(* IEC 61131-3 sources: JingjiangArm/moonboxpro_arm_8.4/Application/Application/任务列表/TensionTask/电机运动/MotionCtl_Gear/PrnVelCtl, 9 files *)

(* ---- KS_CalcMovePara.st ---- *)
(*@CES
Name=KS_CalcMovePara
Type=FunctionBlock
TypeGuid=6f9dac99-8de1-4efc-8465-68ac443b7d08
Guid=11217540-9eff-4725-bda6-b930b9e4eccf
HasDeclaration=True
HasImplementation=True
*)
{DECLARATION}
FUNCTION KS_CalcMovePara : LREAL(*计算运动时间参数|
								控制为even段|只考虑了目标轴匀速、当前轴加速
								返回值作为最终的加速时间s|
								如果时间不能被运动时间间隔整除则会存在pt写入按照整数个
								时间间隔，这里监控的p是使用实际时间的，但是对最终的位置偏差
								没影响。
								负值为返回错误
								-1 参数错误*)
VAR_INPUT
	i_lrVelSa:LREAL;(*启动速度m/min|V0*)
	i_lrVelTar:LREAL;(*目标速度m/min|Vt*)
	i_iDeltime:INT:=21;(*速度规划间隔时间ms|pt运动时间*)
	i_lrGirth_Axis:LREAL;(*轴周长|mm*)
	i_lrReductionRatio:LREAL;(*减速比|电机侧/版辊侧*)
	i_lrDeltPos_Init:LREAL;(*初始位置偏差Pul|开始运动时目标轴和当前轴的位置p偏差*)
	i_lrDeltPos_Final:LREAL;(*最终偏差Pul|最终的目标轴和当前轴的p偏差*)
	i_dwMotorPPR:DWORD:=2097152;(*电机运动一圈的值*)
	i_iSetTime:INT;(*用来计算模数s|*)
END_VAR
VAR
	lrDeltV: LREAL;(*mm/ms*)
	uiTime_N: UINT;(**)
	iDeltT: INT;(*ms*)
	lrCoeff_Axis: LREAL;(*当前轴的比例|Pul/mm*)
	lrRtnValue: LREAL:=0;(*返回值*)
	lrVt: LREAL;(*mm/ms*)
	lrVo: LREAL;(*mm/ms*)
	lrGirth_Axis: LREAL;
	lrDeltPos_Init: LREAL;(*Pul*)
	lrDeltPos_Final:LREAL;(*Pul*)
	(*计算临时变量*)
	uiModCoeff: UINT;(*圈数取整值*)

	lrTemp: LREAL;
	lrTemp1: LREAL;

	(*目标轴位移|mm*)
	lrS_Tar: LREAL;
	(*当前轴位移|mm*)
	lrS_Cur: LREAL;
	dwTime_ms:DWORD;
	lrDelP: LREAL;
	lrDeltS: LREAL;
	lrTime:LREAL;

	lrWatchS_Tar: LREAL;
	lrWatchS_Cur: LREAL;
	lrWatchP_Tar: LREAL;
	lrWatchP_Cur: LREAL;
	lrA: LREAL;
	uiN: UINT;
	iSetTime: INT;
END_VAR
{IMPLEMENTATION}
IF i_lrVelTar<=i_lrVelSa THEN
	lrRtnValue:=-1;
END_IF
lrVt:=i_lrVelTar/60;
lrVo:=i_lrVelSa/60;
lrDeltV:=lrVt-lrVo;

iDeltT:=i_iDeltime;
IF i_iDeltime<=0 THEN
	lrRtnValue:=-1;
END_IF

(*当前轴周长*)
lrGirth_Axis:=i_lrGirth_Axis;
IF lrGirth_Axis<=0 THEN
	lrRtnValue:=-1;
END_IF

IF i_dwMotorPPR<=0 THEN
	lrRtnValue:=-1;
END_IF

IF i_lrReductionRatio<=0 THEN
	lrRtnValue:=-1;
END_IF

(*初始位置偏差Pul|开始运动时目标轴和当前轴的位置p偏差*)
lrDeltPos_Init:=i_lrDeltPos_Init;
lrDeltPos_Init:=KS_MOD_LREAL(lrDeltPos_Init,(i_dwMotorPPR*i_lrReductionRatio));

(*最终偏差Pul|最终的目标轴和当前轴的p偏差*)
lrDeltPos_Final:=i_lrDeltPos_Final;
lrDeltPos_Final:=KS_MOD_LREAL(lrDeltPos_Final,(i_dwMotorPPR*i_lrReductionRatio));

iSetTime:=i_iSetTime;
IF i_iSetTime>=500 THEN(*防止溢出*)
	iSetTime:=500;
END_IF

IF lrRtnValue=0 THEN(*未有错误*)
	dwTime_ms:=(iSetTime)*1000;
	uiTime_N:=(iSetTime)*1000/iDeltT;
	lrA:=lrDeltV/dwTime_ms;

	(*当前轴比例|版辊距离mm转换为电机脉冲值*)
	lrCoeff_Axis:=i_lrReductionRatio*i_dwMotorPPR/i_lrGirth_Axis;(*Pul/mm*)

	(*计算模数值*)
	(*运动的位移*)
	lrS_Tar:=lrVt*dwTime_ms;(*mm*)
	lrS_Cur:=uiTime_N*lrVo*iDeltT+0.5*lrA*iDeltT*iDeltT*uiTime_N*(1+uiTime_N)+
			lrVt*(dwTime_ms-uiTime_N*iDeltT);(*mm*)
	lrDeltS:=lrS_Tar-lrS_Cur;
	IF lrDeltS<=0 THEN
		lrRtnValue:=-2;
	END_IF

	(*转换为电机侧的脉冲*)
	lrDelP:=lrDeltS*lrCoeff_Axis;

	lrTemp:=lrDeltPos_Init+lrDelP-lrDeltPos_Final;
	IF lrTemp<=0 THEN
		lrRtnValue:=-3;
	END_IF
	lrTemp1:=i_dwMotorPPR*i_lrReductionRatio;

	lrTemp:=lrTemp/lrTemp1;
	(*取整数*)

	(*圈数值取整数|版辊圈数*)
	uiModCoeff:=LREAL_TO_UINT(lrTemp);
	IF uiModCoeff<lrTemp THEN
		uiModCoeff:=uiModCoeff+1;
	END_IF

	(*计算需要的时间|按照这个时间可以在目标速度时达到位置同步*)
	IF lrRtnValue=0 THEN
		(*反算时间*)
		lrDelP:=lrDeltPos_Final+uiModCoeff*i_lrReductionRatio*i_dwMotorPPR-lrDeltPos_Init;
		lrDeltS:=lrDelP/lrCoeff_Axis;

		(*寻找复合条件的时间|时间/21的余数小于21*)
		FOR uiN:=uiTime_N TO uiTime_N+10000  BY 1 DO
			lrTemp:=lrDeltV*iDeltT*iDeltT*(1+uiN)*uiN*0.5;
			lrTemp1:=(-lrDeltS-uiN*lrVo*iDeltT+uiN*iDeltT*lrVt);
			lrTime:=lrTemp/lrTemp1;

			IF lrTime-uiN*iDeltT<=iDeltT THEN
				EXIT;
			END_IF

			IF uiN=uiTime_N+10000 THEN(*没有找到|输出负值 标记*)
				lrTime:=-4;
			END_IF
		END_FOR

	END_IF

	IF lrRtnValue=0 THEN
		lrRtnValue:=LREAL_TO_REAL(lrTime/1000);

		(*用于监控*)
		lrWatchS_Tar:=lrVt*lrTime;(*mm*)
		uiTime_N:=uiN;
		lrA:=lrDeltV/lrTime;
		lrWatchS_Cur:=uiTime_N*lrVo*iDeltT+0.5*lrA*iDeltT*iDeltT*uiTime_N*(1+uiTime_N)+
					lrVt*(lrTime-uiTime_N*iDeltT);(*mm*)
		lrWatchP_Tar:=lrWatchS_Tar*lrCoeff_Axis;
		lrWatchP_Cur:=lrWatchS_Cur*lrCoeff_Axis;
	END_IF
END_IF
KS_CalcMovePara:=lrRtnValue;

(* ---- KS_GetInitSts.st ---- *)
(*@CES
Name=KS_GetInitSts
Type=FunctionBlock
TypeGuid=6f9dac99-8de1-4efc-8465-68ac443b7d08
Guid=7ae6f696-fe0b-48ae-942d-bfb0aac909fe
HasDeclaration=True
HasImplementation=True
*)
{DECLARATION}
FUNCTION KS_GetInitSts : BYTE(*获取初始值状态|返回修改的状态*)
VAR_INPUT
	i_bySwitchType:BYTE;(*切换方式|0-空转状态下不考虑单联动状态下都可以切换运动状态
								  |1-空转状态下只有处于联动状态下的轴可以切换*)
	i_xLinkageKnob: BOOL;(*联动旋钮*)
	i_xLinkageSts: BOOL;(*联动状态*)
END_VAR
VAR
	byAxisMotionSts: BYTE;
END_VAR
{IMPLEMENTATION}
IF i_bySwitchType=0 THEN(*空转状态下不考虑单联动状态下都可以切换运动状态*)
	IF i_xLinkageKnob THEN
		byAxisMotionSts:= 0;
	ELSE
		byAxisMotionSts:= 2;
	END_IF
ELSIF i_bySwitchType=1 THEN(*空转状态下只有处于联动状态下的轴可以切换*)
	IF i_xLinkageSts THEN
		byAxisMotionSts:=0;
	ELSE
		byAxisMotionSts:=2;
	END_IF
END_IF
KS_GetInitSts:=byAxisMotionSts;

(* ---- KS_GetMotionSts.st ---- *)
(*@CES
Name=KS_GetMotionSts
Type=FunctionBlock
TypeGuid=6f9dac99-8de1-4efc-8465-68ac443b7d08
Guid=c01ac71d-e678-459d-bed7-b9a659b9ae68
HasDeclaration=True
HasImplementation=True
*)
{DECLARATION}
FUNCTION KS_GetMotionSts : BOOL(*色组轴的运动状态处理|只在开机时候使用 同时控制压辊合压状态|Liu.yt
										轴运动状态标志|0:同步运动状态.
													  |1:同步运动时停止运动状态.
													  |2:停止运动状态
													  |3:停止运动时加速到单运行速度状态.
													  |4:单运行时减速到停止状态.
													  |5:停止运动时或者使用单运行速度运行时加速到同步运动状态.
													  |6:非同步运动时急停到0状态.
													  |7:非同步运动时空转停机到0状态.*)
(*2022.9.21.154927 6,7步中停止的条件判断写错了*)
(*2022.11.29.232720 轴速度是带方向|作为条件需要增加取绝对值*)
(*2023.11.27.165212 增加印刷是否能切换单联动的选择输入接口*)
VAR_INPUT
	i_iGrpId: INT;
	i_xMotionStsSwitchEn:BOOL;(*切换使能|使用该功能需要常有效*)
	i_bySwitchType:BYTE;(*切换方式|0-空转状态下不考虑单联动状态下都可以切换运动状态
								  |1-空转状态下只有处于联动状态下的轴可以切换*)
	i_iGrpAxisNum_Pu: INT; (*色组轴数量*)
	i_pstStSysParam: POINTER TO StSysParam;
//	i_pstStGrpParam: POINTER TO StGrpParam;(*系参数访问入口|*)
	i_paiGrpAxisList: POINTER TO ARRAY [1..MAX_STATION_NUM] OF INT; (*系内所有轴的列表*)
//	i_pastStAxisParam: POINTER TO ARRAY [1..MAX_STATION_NUM] OF StAxisParam;
	i_pastStIOMap_Main_FE						: POINTER TO ARRAY [1..4] OF StIOMap_Main_FE;(*轴io数据区域|AB系*)
	i_pastStIOMap_Axis_FE					: POINTER TO ARRAY [1..MAX_UNIT_NUM] OF StIOMap_Axis_FE;(*轴io数据区域|`````````````````````````````````````````````*)
//	i_pastStIOMap_AxisBasic: POINTER TO ARRAY [1..MAX_STATION_NUM] OF StIOMap_AxisBasic;(*基础io映射表|*)
	i_pabyAxisMotionSts: POINTER TO ARRAY [1..MAX_STATION_NUM] OF BYTE;(*轴运动状态|*)
	i_paxAxisInching:POINTER TO ARRAY [1..MAX_STATION_NUM] OF BOOL;(*轴在单运行|用于控制单运行指示灯显示*)
	i_paxLastAxisInchBtn:POINTER TO ARRAY [1..MAX_STATION_NUM] OF BOOL;(*轴的单运行按钮保留值|用于判断沿*)
	i_iMaxVel_StsSwitch:INT;(*状态切换的最大速度*)
	i_pxFlag_StsSwitchEn:POINTER TO BOOL;(*状态切换使能标志@内部的状态切换标志*)
	i_xChangLinkageStsWhenPrint:BOOL;(*印刷时候可以切换单联动@2023.11.27.164606*)
END_VAR
VAR

	iN: INT;
	xFlag_StsSwitchEn: BOOL;(*状态切换标志*)
	xStsSwitchEn: BOOL;(*状态切换使能*)
	xRetainStsEn: BOOL;(*保持状态标志*)
	iUnitId: INT;
	byAxisMotionSts: BYTE;
	xLastAxisInchBtn: BOOL;
	xAxisInching: BOOL;
	pstStUnitParam_Save: POINTER TO StUnitParam_Save;
	pstStUnitParam_UnSave: POINTER TO StUnitParam_UnSave;
	pstStGrpParam_Save: POINTER TO StGrpParam_Save;
	pstStGrpParam_UnSave: POINTER TO StGrpParam_UnSave;
	pstStIOMap_Axis_FE: POINTER TO StIOMap_Axis_FE;
	xCanSwitchSts_CurAxis: BOOL;(*当前轴可以切换状态标志*)
	dwAxisMotionStsNotOk: DWORD;
END_VAR
{IMPLEMENTATION}
IF i_pstStSysParam<>0 AND
	i_paiGrpAxisList<>0 AND
	i_pastStIOMap_Main_FE<>0 AND
	i_pastStIOMap_Axis_FE<>0 AND
	i_pabyAxisMotionSts<>0 AND
	i_paxAxisInching<>0 AND
	i_paxLastAxisInchBtn<>0 AND
	i_iGrpAxisNum_Pu>0 AND
	i_pxFlag_StsSwitchEn<>0 THEN(*参数合法*)

	xFlag_StsSwitchEn:=i_pxFlag_StsSwitchEn^;
	pstStGrpParam_Save:= ADR(i_pstStSysParam^.astStGrpParam_Save[i_iGrpId]);
	pstStGrpParam_UnSave:= ADR(i_pstStSysParam^.astStGrpParam_UnSave[i_iGrpId]);
	(*2023.11.27.171042 增加了印刷时候有单联动切换的选择接口*)
	xStsSwitchEn:= (pstStGrpParam_UnSave^.xFlag_Ink OR(*空转状态下可以使用|*)
					(pstStGrpParam_UnSave^.xFlag_Print AND i_xChangLinkageStsWhenPrint)) AND
					pstStGrpParam_UnSave^.rVel_Cur<=i_iMaxVel_StsSwitch;(*小于速度限制可以使用*)
	(*印刷时候或者超过限制速度时候|与xStsSwitchEn搭配使用*)
	xRetainStsEn:=(pstStGrpParam_UnSave^.xFlag_Print AND NOT i_xChangLinkageStsWhenPrint)
				OR pstStGrpParam_UnSave^.rVel_Cur>i_iMaxVel_StsSwitch;

	(*切换条件处理*)
	IF  xStsSwitchEn THEN
		xFlag_StsSwitchEn:=TRUE;
	END_IF

	IF i_xMotionStsSwitchEn THEN
		FOR iN:=1 TO i_iGrpAxisNum_Pu BY 1 DO
			iUnitId:=i_paiGrpAxisList^[iN];
			pstStUnitParam_Save:=ADR(i_pstStSysParam^.astStUnitParam_Save[iUnitId]);
			pstStUnitParam_UnSave:=ADR(i_pstStSysParam^.astStUnitParam_UnSave[iUnitId]);
			pstStIOMap_Axis_FE:=ADR(i_pastStIOMap_Axis_FE^[iUnitId]);
			byAxisMotionSts:=i_pabyAxisMotionSts^[iUnitId];
			xLastAxisInchBtn:=i_paxLastAxisInchBtn^[iUnitId];
			xAxisInching:=i_paxAxisInching^[iUnitId];

			xCanSwitchSts_CurAxis:=FALSE;
			IF i_bySwitchType=0 THEN(*空转状态下不考虑单联动状态下都可以切换运动状态*)
				xCanSwitchSts_CurAxis:= pstStUnitParam_UnSave^.xMoveEnable_Motor;
			ELSIF i_bySwitchType=1 THEN(*空转状态下只有处于联动状态下的轴可以切换*)
				xCanSwitchSts_CurAxis:= pstStUnitParam_Save^.xLinkage;
			END_IF

			IF xCanSwitchSts_CurAxis THEN
				CASE byAxisMotionSts OF
					0:(*同步运动状态|此时检查但联动旋钮的状态*)
						IF NOT pstStIOMap_Axis_FE^.i_xLinkage AND (*切换到单动状态*)
							NOT pstStIOMap_Axis_FE^.o_xRel_Press THEN(*压辊未合压时起作用*)
							byAxisMotionSts:=1;
						END_IF
					1:(*处于停止运动过程状态|等待到达停止运动状态*)
						IF pstStIOMap_Axis_FE^.i_xLinkage THEN(*联动状态|恢复到同步运动状态*)
							byAxisMotionSts:=5;
						END_IF

						IF byAxisMotionSts=1 THEN
							IF ABS(pstStUnitParam_UnSave^.rAxisVel_PrnRoller)<=0.0001 THEN(*减速到0我们认为到达了停止运动状态*)
								byAxisMotionSts:=2;
							END_IF
						END_IF
					2:(*停止运动状态*)
						IF pstStIOMap_Axis_FE^.i_xLinkage THEN(*联动状态|恢复到同步运动状态*)
							byAxisMotionSts:=5;
						END_IF

						(*检查单运行是否按下*)
						IF byAxisMotionSts=2 THEN
							IF pstStIOMap_Axis_FE^.i_xInch AND NOT xLastAxisInchBtn THEN(*单运行按下了*)
								byAxisMotionSts:=3;
							END_IF
						END_IF

					3:(*加速到单运行状态*)
						IF pstStIOMap_Axis_FE^.i_xLinkage THEN(*联动状态|恢复到同步运动状态*)
							byAxisMotionSts:=5;
						END_IF

						IF byAxisMotionSts=3 THEN
							IF (pstStIOMap_Axis_FE^.i_xInch AND NOT xLastAxisInchBtn) OR(*单运行按下了*)
								NOT xStsSwitchEn THEN(*退出了状态*)
								byAxisMotionSts:=4;
							END_IF
						END_IF
					4:(*单运行状态停止到停止状态*)
						IF pstStIOMap_Axis_FE^.i_xLinkage THEN(*联动状态|恢复到同步运动状态*)
							byAxisMotionSts:=5;
						END_IF

						IF byAxisMotionSts=4 THEN
							IF ABS(pstStUnitParam_UnSave^.rAxisVel_PrnRoller)<=0.0001 THEN(*减速到0我们认为到达了停止运动状态*)
								byAxisMotionSts:=2;
							END_IF
						END_IF
					5:(*前往同步运动状态*)
						IF NOT pstStIOMap_Axis_FE^.i_xLinkage THEN(*切换到单动状态*)
							byAxisMotionSts:=1;
						END_IF

						IF byAxisMotionSts=5 THEN
							IF ABS(ABS(pstStUnitParam_UnSave^.rAxisVel_PrnRoller)-pstStGrpParam_UnSave^.rVel_Cur)<=0.0001 THEN(*到达当前速度*)
								byAxisMotionSts:=0;
							END_IF
						END_IF
					6,7:(*非同步状态下非停止状态下的停止和急停*)
						IF ABS(pstStUnitParam_UnSave^.rAxisVel_PrnRoller)<=0.0001 THEN(*到达0速度|2022.9.21.154723 -以前的条件写错了*)
							byAxisMotionSts:=KS_GetInitSts(i_bySwitchType,
													pstStIOMap_Axis_FE^.i_xLinkage,
													pstStUnitParam_Save^.xLinkage);
						END_IF
				ELSE
					byAxisMotionSts:=KS_GetInitSts(i_bySwitchType,
											pstStIOMap_Axis_FE^.i_xLinkage,
											pstStUnitParam_Save^.xLinkage);
				END_CASE
			ELSE
				byAxisMotionSts:=KS_GetInitSts(i_bySwitchType,
										pstStIOMap_Axis_FE^.i_xLinkage,
										pstStUnitParam_Save^.xLinkage);
			END_IF

			(*处理单运行指示*)
			IF byAxisMotionSts=3 OR(*单运行加速*)
				byAxisMotionSts=4 THEN(*单运行减速*)
				xAxisInching:=TRUE;
			ELSE
				xAxisInching:=FALSE;
			END_IF

			(*切换使能无效了-在状态恢复到初始状态时候xFlag_StsSwitchEn标志为false|
			byAxisMotionSts 在停机时候强制写为初值|
							在印刷状态或者超过限制速度时不切换|*)
			IF xRetainStsEn THEN(*保持之前状态|*)
				byAxisMotionSts:=i_pabyAxisMotionSts^[iUnitId];
			ELSE
				IF NOT xFlag_StsSwitchEn THEN
					byAxisMotionSts:=KS_GetInitSts(i_bySwitchType,
												pstStIOMap_Axis_FE^.i_xLinkage,
												pstStUnitParam_Save^.xLinkage);
				END_IF
			END_IF

			(*处理停机和急停*)
			IF byAxisMotionSts<>0 AND  byAxisMotionSts<>2 THEN
				IF pstStGrpParam_UnSave^.xFlag_EStoping THEN(*急停过程中|*)
					byAxisMotionSts:=6;
				ELSIF pstStGrpParam_UnSave^.xFlag_Ink AND
					(pstStGrpParam_UnSave^.xFlag_Stoping OR (*空转停止过程中*)
					pstStGrpParam_UnSave^.xFlag_FastStoping) THEN
					byAxisMotionSts:=7;
				END_IF

				(*判断轴运动状态|未处于停止状态或者同步状态|*)
				dwAxisMotionStsNotOk:=dwAxisMotionStsNotOk OR SHL(DWORD#1,iUnitId-1);
			END_IF

			(*使能模式控制|2022.7.14.121739*)
			IF i_bySwitchType=0 THEN
				IF byAxisMotionSts=2 THEN(*停止状态 写3*)
					pstStUnitParam_Save^.wEnableMode_Motor:=3;
				ELSE(*非停止状态|写4*)
					pstStUnitParam_Save^.wEnableMode_Motor:=4;
				END_IF
			ELSE
				IF pstStUnitParam_Save^.wEnableMode_Motor=3 OR
					pstStUnitParam_Save^.wEnableMode_Motor=4 THEN(*说明进行过使能切换|此时强制将使能模式写成4*)
					pstStUnitParam_Save^.wEnableMode_Motor:=4;
				ELSE
					pstStUnitParam_Save^.wEnableMode_Motor:=0;
				END_IF
			END_IF

			i_pabyAxisMotionSts^[iUnitId]:=byAxisMotionSts;
			i_paxAxisInching^[iUnitId]:=xAxisInching;
			i_paxLastAxisInchBtn^[iUnitId]:=i_pastStIOMap_Axis_FE^[iUnitId].i_xInch;
		END_FOR

		(*切换条件处理*)
		IF NOT xStsSwitchEn THEN
			IF xFlag_StsSwitchEn THEN
				IF dwAxisMotionStsNotOk=0 THEN(*都处于初始态|可以清除标志了*)
					xFlag_StsSwitchEn:=FALSE;
				END_IF
			END_IF
		END_IF
	ELSE(*不使能*)
		FOR iN:=1 TO i_iGrpAxisNum_Pu BY 1 DO
			iUnitId:=i_paiGrpAxisList^[iN];
			pstStUnitParam_Save:=ADR(i_pstStSysParam^.astStUnitParam_Save[iUnitId]);
			pstStUnitParam_UnSave:=ADR(i_pstStSysParam^.astStUnitParam_UnSave[iUnitId]);
			i_pabyAxisMotionSts^[iUnitId]:=0;
			i_paxAxisInching^[iUnitId]:=FALSE;
			i_paxLastAxisInchBtn^[iUnitId]:=FALSE;

			IF pstStUnitParam_Save^.wEnableMode_Motor=3 OR
				pstStUnitParam_Save^.wEnableMode_Motor=4 THEN(*说明进行过使能切换|此时强制将使能模式写成4*)
				pstStUnitParam_Save^.wEnableMode_Motor:=4;
			ELSE
				pstStUnitParam_Save^.wEnableMode_Motor:=0;
			END_IF
		END_FOR
		xFlag_StsSwitchEn:=FALSE;
	END_IF

	i_pxFlag_StsSwitchEn^:=xFlag_StsSwitchEn;
END_IF

(* ---- KS_GetRelatePos.st ---- *)
(*@CES
Name=KS_GetRelatePos
Type=FunctionBlock
TypeGuid=6f9dac99-8de1-4efc-8465-68ac443b7d08
Guid=64bf2139-19b0-44f0-86e4-ed0fdab8fbfc
HasDeclaration=True
HasImplementation=True
*)
{DECLARATION}
FUNCTION KS_GetRelatePos : BOOL(*计算所有目标轴和当前轴的相对位置|节省空间就只做16个轴
								目标轴为联动非涂布轴*)
VAR_INPUT
	i_iAxisId_Cur:INT;(*当前轴id*)
	i_iGrpAxisNum_Pu: INT; (*色组轴数量*)
	i_paiGrpAxisList: POINTER TO ARRAY [1..MAX_UNIT_NUM] OF INT; (*系内所有轴的列表*)
	i_pastStUnitParam_Save: POINTER TO ARRAY [1..MAX_UNIT_NUM] OF StUnitParam_Save;
	i_pastStUnitParam_UnSave: POINTER TO ARRAY [1..MAX_UNIT_NUM] OF StUnitParam_UnSave;
	i_palrRelatePos:POINTER TO ARRAY [1..MAX_UNIT_NUM] OF LREAL;(*索引为目标轴*)
END_VAR
VAR
	in: INT;
	iAxisId: INT;
	pstStUnitParam_Save: POINTER TO StUnitParam_Save;
	pstStUnitParam_UnSave: POINTER TO StUnitParam_UnSave;
	pstStUnitParam_Cur_UnSave: POINTER TO StUnitParam_UnSave;
	ailist: ARRAY [1..MAX_STATION_NUM] OF INT;(*联动非涂布列表|不包含当前色*)
	iIndex:INT;
	xDne: BOOL;(*获取成功了*)
END_VAR
{IMPLEMENTATION}
(*初始化*)
IF	i_palrRelatePos<>0	THEN
	FOR iN:=1 TO 16 BY 1 DO
		i_palrRelatePos^[iN]:=0;
	END_FOR
END_IF
iIndex:=0;
IF i_iAxisId_Cur>0 AND
	i_iAxisId_Cur<=16 AND
	i_iGrpAxisNum_Pu>1 AND
	i_paiGrpAxisList<>0 THEN
	pstStUnitParam_Cur_UnSave:=ADR(i_pastStUnitParam_UnSave^[i_iAxisId_Cur]);
	FOR in:=1 TO i_iGrpAxisNum_Pu BY 1 DO
		iAxisId:=i_paiGrpAxisList^[iN];
		IF iAxisId<>i_iAxisId_Cur THEN(*非当前轴*)
			pstStUnitParam_Save:=ADR(i_pastStUnitParam_Save^[iAxisId]);
			IF pstStUnitParam_Save^.xLinkage AND(*联动*)
				NOT pstStUnitParam_Save^.xSwitchOn_CoatingPrn THEN(*非涂布色组*)
				iIndex:=iIndex+1;
				ailist[iIndex]:=iAxisId;
			END_IF
		END_IF
	END_FOR

	FOR iN:=1 TO iIndex BY 1 DO
		iAxisId:=ailist[iN];
		pstStUnitParam_UnSave:=ADR(i_pastStUnitParam_UnSave^[iAxisId]);
		i_palrRelatePos^[iAxisId]:=pstStUnitParam_UnSave^.lrPrf_Pos-pstStUnitParam_Cur_UnSave^.lrPrf_Pos;
		xDne:=TRUE;
	END_FOR
END_IF
KS_GetRelatePos:=xDne;

(* ---- KS_GetUnitId_Tar.st ---- *)
(*@CES
Name=KS_GetUnitId_Tar
Type=FunctionBlock
TypeGuid=6f9dac99-8de1-4efc-8465-68ac443b7d08
Guid=50ffccd4-38ae-4948-a424-e85895436bf8
HasDeclaration=True
HasImplementation=True
*)
{DECLARATION}
FUNCTION KS_GetUnitId_Tar : INT(*获取目标轴id|轴号1--16*)
VAR_INPUT
	i_iUnitId_Cur:INT;(*当前轴id*)
	i_iGrpAxisNum_Pu: INT; (*色组轴数量*)
	i_paiGrpAxisList: POINTER TO ARRAY [1..MAX_STATION_NUM] OF INT; (*系内所有轴的列表*)
	i_pastStUnitParam_Save: POINTER TO ARRAY [1..MAX_UNIT_NUM] OF StUnitParam_Save;
	i_pastStUnitParam_UnSave: POINTER TO ARRAY [1..MAX_UNIT_NUM] OF StUnitParam_UnSave;
	i_pabyAxisMotionSts: POINTER TO ARRAY [1..MAX_STATION_NUM] OF BYTE;(*轴运动状态|*)
END_VAR
VAR
	iUnitId_Tar: INT;
	iUnitId:INT;
	pstStUnitParam_Save: POINTER TO StUnitParam_Save;
	pstStUnitParam_UnSave: POINTER TO StUnitParam_UnSave;
	iN: INT;
END_VAR
{IMPLEMENTATION}
iUnitId_Tar:=-1;
IF i_iUnitId_Cur>0 AND
	i_iUnitId_Cur<=16 AND
	i_iGrpAxisNum_Pu>1 AND
	i_paiGrpAxisList<>0 AND
	i_pastStUnitParam_Save<>0 AND
	i_pastStUnitParam_UnSave<>0 AND
	i_pabyAxisMotionSts<>0 THEN

	FOR iN:=1 TO i_iGrpAxisNum_Pu BY 1 DO
		iUnitId:=i_paiGrpAxisList^[iN];
		IF iUnitId<>i_iUnitId_Cur THEN
			pstStUnitParam_Save:=ADR(i_pastStUnitParam_Save^[iUnitid]);

			IF pstStUnitParam_Save^.xLinkage AND(*联动*)
				NOT pstStUnitParam_Save^.xSwitchOn_CoatingPrn AND(*非涂布色组*)
				i_pabyAxisMotionSts^[iUnitId]=0 THEN(*处于同步运动状态*)
				iUnitId_Tar:=iUnitId;
				EXIT;
			END_IF
		END_IF
	END_FOR
END_IF
KS_GetUnitId_Tar:=iUnitId_Tar;

(* ---- KS_VelPrfByAxisMotionSts.st ---- *)
(*@CES
Name=KS_VelPrfByAxisMotionSts
Type=FunctionBlock
TypeGuid=6f9dac99-8de1-4efc-8465-68ac443b7d08
Guid=bab22195-914f-4e07-a531-52e1aa67a074
HasDeclaration=True
HasImplementation=True
*)
{DECLARATION}
FUNCTION KS_VelPrfByAxisMotionSts : BOOL(*根据轴运动状态标志控制轴速度输出
													  |0:同步运动状态.
													  |1:同步运动时停止运动状态.
													  |2:停止运动状态
													  |3:停止运动时加速到单运行速度状态.
													  |4:单运行时减速到停止状态.
													  |5:停止运动时或者使用单运行速度运行时加速到同步运动状态.
													  |6:非同步运动时急停到0状态.
													  |7:非同步运动时空转停机到0状态.*)
(*该功能的加减速时间分开|2022.5.29.004252*)
(*2022.12.26.135440 |出现过因为pstStAxisParam^.byEnableModeSwitchDne.1变量作为速度规划条件的时候
因为停机时机的问题引起的速度不能清除的问题，使用本地变量作为条件*)
(*2023.2.15.173943 所有的减速时间都由手动减速时间修改为了停止时间*)
(*2023.07.24.171926处理因为时序问题引起的motionctl中不能正确设置当前伺服状态*)
VAR_INPUT
	i_iGrpId: INT;
	i_iGrpAxisNum_Pu: INT; (*色组轴数量*)
	i_pstStSysParam: POINTER TO StSysParam;
//	i_pstStGrpParam: POINTER TO StGrpParam;(*系参数访问入口|*)
	i_paiGrpAxisList: POINTER TO ARRAY [1..MAX_UNIT_NUM] OF INT; (*系内所有轴的列表*)
//	i_pastStAxisParam: POINTER TO ARRAY [1..MAX_STATION_NUM] OF StAxisParam;
	i_pabyAxisMotionSts: POINTER TO ARRAY [1..MAX_STATION_NUM] OF BYTE;(*轴运动状态*)
	i_palrAxisMotionVel:POINTER TO ARRAY [1..MAX_STATION_NUM] OF LREAL;(*轴速度*)
	i_palrAcceleToSync:POINTER TO ARRAY [1..16] OF LREAL;(*用来保证同步的加速度|m/min/ms|16个轴*)
	i_xMotionEnabled: BOOL;(*MotionCtl功能块准备好了|可以规划速度|2022.7.14.133144*)
	i_pxVelPrfEn: POINTER TO BOOL;(*可以规划速度已经使能|2022.7.14.133144*)
	i_xNeedKeepSync:BOOL;(*需要保证同步|在前往同步时候如果加减速有效了-则按照界面输入时间进行加减速|2022.7.21.174859*)
	i_paxAxisVelPrfEn:POINTER TO ARRAY [1..MAX_STATION_NUM] OF BOOL;(*2022.12.26.135324 增加了轴速度的规划使能标志|进行速度规划的条件*)
	i_uiMaxVel_UseCalcAcc:UINT;(*用于计算最大加速度的最大速度@2024.04.12.180552*)
END_VAR
VAR
	iTimeAccDec: INT;(*加减速时间|s|正负标记加减速*)
	lrVel_Max: REAL;(*最大速度*)
	lrDelVelPerCycle: LREAL;(*单位周期的速度变化*)
	pstStUnitParam_Save: POINTER TO StUnitParam_Save;
	pstStUnitParam_UnSave: POINTER TO StUnitParam_UnSave;
	abyLastAxisMotionSts:ARRAY [1..MAX_STATION_NUM] OF BYTE;
	iN: INT;
	iUnitId: INT;
	byAxisMotionSts: BYTE;
	byLastAxisMotionSts: BYTE;
	lrAxisMotionVel: LREAL;
	lrVel_Cur: LREAL;
	lrVel_Tar: LREAL;
	xUseInputAccele: BOOL;(**)
	dwAxisVelPrfMustEnable: DWORD;
END_VAR
{IMPLEMENTATION}
IF i_pstStSysParam<>0 AND
	i_paiGrpAxisList<>0 AND
	i_pabyAxisMotionSts<>0 AND
	i_iGrpAxisNum_Pu>0 AND
	i_palrAxisMotionVel<>0 AND
	i_palrAcceleToSync<>0 AND
	i_pxVelPrfEn<>0 AND
	i_paxAxisVelPrfEn<>0 THEN

	IF i_xMotionEnabled  THEN(*上伺服模式写为4成功后执行速度控制*)
		i_pxVelPrfEn^:=TRUE;
	END_IF

	FOR iN:=1 TO i_iGrpAxisNum_Pu BY 1 DO
		iUnitId:=i_paiGrpAxisList^[iN];
		byAxisMotionSts:=i_pabyAxisMotionSts^[iUnitId];
		byLastAxisMotionSts:=abyLastAxisMotionSts[iUnitId];
		lrAxisMotionVel:=i_palrAxisMotionVel^[iUnitId];
		pstStUnitParam_Save:=ADR(i_pstStSysParam^.astStUnitParam_Save[iUnitId]);
		pstStUnitParam_UnSave:=ADR(i_pstStSysParam^.astStUnitParam_UnSave[iUnitId]);

		(*2023.07.24.171926@将清除位置移动到此处|
		处理因为时序问题引起的motionctl中不能正确设置当前伺服状态*)
		(*2022.12.26.135650@解决异常速度规划不能到0问题*)
		IF i_paxAxisVelPrfEn^[iUnitId] AND
			NOT pstStUnitParam_UnSave^.byEnableModeSwitchDne.1 AND
			lrAxisMotionVel<=0.00001 THEN(*速度规划到0了|复位标志*)
			i_paxAxisVelPrfEn^[iUnitId]:=FALSE;
		END_IF

		(*2022.12.26.135440 |出现过因为pstStAxisParam^.byEnableModeSwitchDne.1变量作为速度规划条件的时候
		因为停机时机的问题引起的速度不能清除的问题，使用本地变量作为条件*)
		IF pstStUnitParam_UnSave^.byEnableModeSwitchDne.1 THEN
			i_paxAxisVelPrfEn^[iUnitId]:=pstStUnitParam_UnSave^.byEnableModeSwitchDne.1;
		END_IF

		(*2024.12.31.102049 同步*)
		IF pstStUnitParam_Save^.xSwitchOn_CoatingPrn THEN(*涂布*)
			lrVel_Cur:=pstStUnitParam_UnSave^.lrVelocity_CoatingPrn;
		ELSE
			(*2024.12.22.164428@色组轴*)
			IF NOT i_pstStSysParam^.stStSysParam_Save.xAxisPrfVelEn THEN
				lrVel_Cur:=i_pstStSysParam^.astStGrpParam_UnSave[i_iGrpId].rVel_Cur;
			ELSE
				//2026.5.9.193956这里更新了，不知道有没有问题
				IF i_pstStSysParam^.astStGrpParam_UnSave[i_iGrpId].xFlag_AutoAcc OR
						i_pstStSysParam^.astStGrpParam_UnSave[i_iGrpId].xFlag_AutoDec THEN
					lrVel_Cur:=pstStUnitParam_UnSave^.rAxisPrfVel;
				ELSE
					lrVel_Cur:=i_pstStSysParam^.astStGrpParam_UnSave[i_iGrpId].rVel_Cur;
				END_IF
			END_IF
		END_IF

		xUseInputAccele:=FALSE;

		CASE byAxisMotionSts OF
			0:(*同步转动状态*)
				lrVel_Tar:=lrVel_Cur;
				iTimeAccDec:=0;(*完全跟随*)
			1:(*同步运动状态下减速到停止状态*)
				lrVel_Tar:=0;
(*				iTimeAccDec:=-i_pstStGrpParam^.iTime_ManuDec;(*手动减速时间跟随*)*)
				iTimeAccDec:=-i_pstStSysParam^.astStGrpParam_Save[i_iGrpId].iTime_Stop;(*停止时间跟随@2023.2.15.174049*)
			2:(*停止运动状态*)
				lrVel_Tar:=0;
(*				iTimeAccDec:=-i_pstStGrpParam^.iTime_ManuDec;(*手动减速时间跟随*)*)
				iTimeAccDec:=-i_pstStSysParam^.astStGrpParam_Save[i_iGrpId].iTime_Stop;(*停止时间跟随@2023.2.15.174049*)
			3:(*停止运动状态加速到单运行速度*)
				lrVel_Tar:=i_pstStSysParam^.astStGrpParam_Save[i_iGrpId].rVel_Inch;
				iTimeAccDec:=i_pstStSysParam^.astStGrpParam_Save[i_iGrpId].iTime_ManuAcc;(*手动加速时间跟随*)
			4:(*单运行减速到停止位置*)
				lrVel_Tar:=0;
(*				iTimeAccDec:=-i_pstStGrpParam^.iTime_ManuDec;(*手动减速时间跟随*)*)
				iTimeAccDec:=-i_pstStSysParam^.astStGrpParam_Save[i_iGrpId].iTime_Stop;(*停止时间跟随@2023.2.15.174049*)
			5:(*加速到同步速度状态*)
				lrVel_Tar:=lrVel_Cur;
				IF lrAxisMotionVel<=lrVel_Tar THEN(*2022.12.26.134601 +条件*)
					iTimeAccDec:=i_pstStSysParam^.astStGrpParam_Save[i_iGrpId].iTime_ManuAcc;(*手动加速时间跟随*)
				ELSE(*2022.12.26.134601 +条件*)
					iTimeAccDec:=-i_pstStSysParam^.astStGrpParam_Save[i_iGrpId].iTime_ManuAcc;(*手动减速时间跟随*)
				END_IF
				IF i_palrAcceleToSync^[iUnitId]<>0 THEN(*说明计算出来了同步*)
					xUseInputAccele:=TRUE;
				END_IF
			6:(*非同步状态时急停到0状态*)
				lrVel_Tar:=0;
				iTimeAccDec:=-i_pstStSysParam^.astStGrpParam_Save[i_iGrpId].iTime_Estop;(*急停时间跟随*)

			7:
				lrVel_Tar:=0;
				iTimeAccDec:=-i_pstStSysParam^.astStGrpParam_Save[i_iGrpId].iTime_stop;(*停止时间跟随*)
		ELSE
			lrVel_Tar:=0;
			iTimeAccDec:=-i_pstStSysParam^.astStGrpParam_Save[i_iGrpId].iTime_Estop;(*急停时间跟随*)
		END_CASE;

		(*速度控制*)
		(*计算加减加速度值*)
		lrVel_Max:=(i_uiMaxVel_UseCalcAcc);
		IF lrVel_Max<=20 THEN(*最大速度限制到20m/min以上*)
			lrVel_Max:=20;
		END_IF
		IF iTimeAccDec<>0 THEN
			lrDelVelPerCycle:=lrVel_Max*gc_iCycleTime_Motion/iTimeAccDec/1000;
			(*由外部计算出的加速度控制到达同步速度时保证位置同步|2021.1.5.155658*)
			IF xUseInputAccele AND i_xNeedKeepSync THEN(*需要使用外部输入的加速度进行加速|2022.7.21.175130增加需要同步使能*)
				lrDelVelPerCycle:=i_palrAcceleToSync^[iUnitId]*gc_iCycleTime_Motion;
			END_IF
			IF i_pxVelPrfEn^ AND
				//NOT i_pstStGrpParam^.xFlag_PTfifofull AND
(*				pstStAxisParam^.byEnableModeSwitchDne.1 THEN*)
				i_paxAxisVelPrfEn^[iUnitId] THEN(*2022.12.26.152739 替换*)

				lrAxisMotionVel:=lrAxisMotionVel+lrDelVelPerCycle;
				IF lrDelVelPerCycle>0 THEN(*加速*)
					IF lrAxisMotionVel>=lrVel_Tar THEN
						lrAxisMotionVel:=lrVel_Tar;
					END_IF
				ELSE(*减速*)
					IF lrAxisMotionVel<=lrVel_Tar THEN
						lrAxisMotionVel:=lrVel_Tar;
					END_IF
				END_IF
			END_IF
		ELSE
			lrAxisMotionVel:=lrVel_Tar;
		END_IF

		IF NOT pstStUnitParam_UnSave^.xMoveEnable_Motor OR(*2022.7.14.102148 联动标志修改为了电机运动使能标志*)
			lrAxisMotionVel<0.00001 THEN(*防止因为数据类型的原因导致值不能完全=0*)
			lrAxisMotionVel:=0.0;
		END_IF

		IF lrAxisMotionVel<>0 THEN(*速度未到0了*)
			dwAxisVelPrfMustEnable:=dwAxisVelPrfMustEnable OR
									SHL(DWORD#1,iUnitId-1);

		END_IF

		i_palrAxisMotionVel^[iUnitId]:=lrAxisMotionVel;
		(*2023.07.24.171926@将清除位置移动到规划使能的位置|
		处理因为时序问题引起的motionctl中不能正确设置当前伺服状态*)
(*
		(*2022.12.26.135650@解决异常速度规划不能到0问题*)
		IF i_paxAxisVelPrfEn^[iAxisId] AND
			NOT pstStAxisParam^.byEnableModeSwitchDne.1 AND
			lrAxisMotionVel<=0.00001 THEN(*速度规划到0了|复位标志*)
			i_paxAxisVelPrfEn^[iAxisId]:=FALSE;
		END_IF
*)
	END_FOR

	(*2022.7.14.134141  *)
	IF i_pxVelPrfEn^ AND
		(NOT i_xMotionEnabled) THEN
		IF dwAxisVelPrfMustEnable=0 THEN(*不需要使能了*)
			i_pxVelPrfEn^:=FALSE;
		END_IF
	END_IF
ELSE;
END_IF

(* ---- KS_FB_AxisVelCtl_PrnRoller.st ---- *)
(*@CES
Name=KS_FB_AxisVelCtl_PrnRoller
Type=FunctionBlock
TypeGuid=6f9dac99-8de1-4efc-8465-68ac443b7d08
Guid=abdd25c9-7f8b-492e-b7cd-5839eca90f4a
HasDeclaration=True
HasImplementation=True
*)
{DECLARATION}
FUNCTION_BLOCK KS_FB_AxisVelCtl_PrnRoller(*色组轴速度控制*)
(*在原来的联动状态下切换单联动状态并保持同步逻辑的基础上
兼容随时单联动切换的速度处理|目前只处理色组轴-2022.7.11.111134*)
VAR_INPUT
	i_xEn:BOOL;
	i_iGrpId: INT;
	i_xSwitchType0:BOOL;(*切换方式|TRUE：空转时候可以随时切换单联动轴的运动状态*)
	i_xSwitchType1:BOOL;(*切换方式|TRUE：空转状态下只能切换已经联动轴的运动状态|
						通过单联动旋钮处理，并能保证切换后相位能够保持之前状态*)
	i_xMotionStsSwitchEn:BOOL;(*切换使能*)
	i_xNeedKeepSync:BOOL;(*需要保证同步|在前往同步时候如果加减速有效了-则按照界面输入时间进行加减速|2022.7.21.174859*)
	i_iGrpAxisNum_Pu: INT; (*色组轴数量*)
	i_pstStSysParam: POINTER TO StSysParam;
//	i_pstStGrpParam: POINTER TO StGrpParam;(*系参数访问入口|*)
	i_paiGrpAxisList: POINTER TO ARRAY [1..MAX_UNIT_NUM] OF INT; (*系内所有轴的列表*)
//	i_pastStAxisParam: POINTER TO ARRAY [1..MAX_STATION_NUM] OF StAxisParam;
	i_pastStIOMap_Main_FE						: POINTER TO ARRAY [1..4] OF StIOMap_Main_FE;(*轴io数据区域|AB系*)
	i_pastStIOMap_Axis_FE					: POINTER TO ARRAY [1..MAX_UNIT_NUM] OF StIOMap_Axis_FE;(*轴io数据区域|`````````````````````````````````````````````*)
//	i_pastStIOMap_AxisBasic: POINTER TO ARRAY [1..MAX_STATION_NUM] OF StIOMap_AxisBasic;(*基础io映射表|*)
	i_pabyAxisMotionSts: POINTER TO ARRAY [1..MAX_UNIT_NUM] OF BYTE;(*轴运动状态|*)
	i_paxAxisInching:POINTER TO ARRAY [1..MAX_UNIT_NUM] OF BOOL;(*轴在单运行|用于控制单运行指示灯显示*)
	i_paxLastAxisInchBtn:POINTER TO ARRAY [1..MAX_UNIT_NUM] OF BOOL;(*轴的单运行按钮保留值|用于判断沿*)
	i_iMaxVel_StsSwitch:INT;(*状态切换的最大速度*)

	i_palrAxisMotionVel:POINTER TO ARRAY [1..MAX_UNIT_NUM] OF LREAL;(*轴速度*)
	i_palrAcceleToSync:POINTER TO ARRAY [1..16] OF LREAL;(*用来保证同步的加速度|m/min/ms|16个轴*)
	i_palrTimeToSync:POINTER TO ARRAY [1..16] OF LREAL;(*同步加到目标速度的时间*)
	i_palrRelatePos_Final:POINTER TO ARRAY [1..16,1..16] OF LREAL;(*做成16个轴|
													记录目标轴和当前轴的相对位置值|最后恢复的位置差
													一维下标为当前轴号，二维下标为目标轴号*)
	i_palrRelatePosToSync:POINTER TO ARRAY [1..16,1..16] OF LREAL;(*做成16个轴|
												记录目标轴和当前轴的相对位置值|开始切换到同步状态时的位置差
												一维下标为当前轴号，二维下标为目标轴号*)
	i_xMotionEnabled: BOOL;(*可以规划速度已经使能|2022.7.14.133144*)
	i_xChangLinkageStsWhenPrint:BOOL;(*印刷时候可以切换单联动@2023.11.27.164606*)
	i_uiMaxVel_UseCalcAcc:UINT;(*用于计算最大加速度的最大速度@2024.04.12.180552*)
END_VAR
VAR_OUTPUT
	o_xEn:BOOL;
END_VAR
VAR
	fbKS_FB_GetAcceleToSync: KS_FB_GetAcceleToSync;
	bySwitchType: BYTE;(*切换方式|0-空转状态下不考虑单联动状态下都可以切换运动状态
								 |1-空转状态下只有处于联动状态下的轴可以切换*)
	xFlag_StsSwitchEn: BOOL;
	xVelPrfEn: BOOL;
	xNeedKeepSync: BOOL;(*需要保证位置同步|在到达同步状态时候*)
	axAxisVelPrfEn: ARRAY [1..MAX_STATION_NUM] OF BOOL;(*2022.12.26.135955+*)
END_VAR
{IMPLEMENTATION}
(*2020.12.24.145952 增加的开机后可以控制色组轴的运动速度|Liu.yt*)
bySwitchType:=255;
IF i_xSwitchType0 THEN
	bySwitchType:=0;
ELSIF i_xSwitchType1 THEN
	bySwitchType:=1;
END_IF

KS_GetMotionSts(
	i_iGrpId,
	i_xMotionStsSwitchEn AND bySwitchType<>255(*i_xMotionStsSwitchEn*),
	bySwitchType,(*I_bySwitchType*)
	i_iGrpAxisNum_Pu(*i_iGrpAxisNum_Pu*),
	i_pstStSysParam,
//i_pstStGrpParam(*i_pstStGrpParam*),
	i_paiGrpAxisList(*i_paiGrpAxisList*),
//	i_pastStAxisParam(*i_pastStAxisParam*),
	i_pastStIOMap_Main_FE,
	i_pastStIOMap_Axis_FE,
//	i_pastStIOMap_AxisBasic(*i_pastStIOMap_AxisBasic*),
	i_pabyAxisMotionSts(*i_pabyAxisMotionSts*),
	i_paxAxisInching(*i_paxAxisInching*),
	i_paxLastAxisInchBtn(*i_paxLastAxisInchBtn*),
	i_iMaxVel_StsSwitch(*i_iMaxVel_StsSwitch*),
	ADR(xFlag_StsSwitchEn)(*i_pxFlag_StsSwitchEn*),
	i_xChangLinkageStsWhenPrint(*i_xChangLinkageStsWhenPrint*));

fbKS_FB_GetAcceleToSync(
	i_xEn:= i_pstStSysParam^.astStGrpParam_UnSave[i_iGrpId].xFlag_Ink ,(*只有空转才能使用*)
	i_iGrpId:= i_iGrpId,
	i_iGrpAxisNum_Pu:= i_iGrpAxisNum_Pu,
	i_pstStSysParam:= i_pstStSysParam,
	i_paiGrpAxisList:= i_paiGrpAxisList,
//	i_pastStAxisParam:= i_pastStAxisParam,
	i_pabyAxisMotionSts:= i_pabyAxisMotionSts,
	i_palrAcceleToSync:=i_palrAcceleToSync,
	i_palrTimeToSync:=i_palrTimeToSync,
	i_palrRelatePos_Final:=i_palrRelatePos_Final,
	i_palrRelatePosToSync:=i_palrRelatePosToSync,
	o_xEn=>);

(**控制速度规划*)
xNeedKeepSync:=i_xNeedKeepSync;
IF i_pstStSysParam^.astStGrpParam_UnSave[i_iGrpId].xFlag_Accing OR
	i_pstStSysParam^.astStGrpParam_UnSave[i_iGrpId].xFlag_Decing THEN
	xNeedKeepSync:=FALSE;(*如果有加速则取消同步*)
END_IF
KS_VelPrfByAxisMotionSts(
	i_iGrpId,
	i_iGrpAxisNum_Pu(*i_iGrpAxisNum_Pu*),
	i_pstStSysParam(*i_pstStGrpParam*),
	i_paiGrpAxisList(*i_paiGrpAxisList*),
//	i_pastStAxisParam(*i_pastStAxisParam*),
	i_pabyAxisMotionSts(*i_pabyAxisMotionSts*),
	i_palrAxisMotionVel(*i_palrAxisMotionVel*),
	i_palrAcceleToSync(*i_palrAcceleToSync*),
	i_xMotionEnabled,
	ADR(xVelPrfEn),
	xNeedKeepSync,
	ADR(axAxisVelPrfEn),
	i_uiMaxVel_UseCalcAcc);

(* ---- KS_FB_Compensate_Vel_Prn.st ---- *)
(*@CES
Name=KS_FB_Compensate_Vel_Prn
Type=FunctionBlock
TypeGuid=6f9dac99-8de1-4efc-8465-68ac443b7d08
Guid=f2c8bddd-aead-4231-9ab2-ee8ef03f3302
HasDeclaration=True
HasImplementation=True
*)
{DECLARATION}
FUNCTION_BLOCK KS_FB_Compensate_Vel_Prn
VAR_INPUT
	i_xEn: BOOL;
	i_iGrpId: INT;
	i_rVel_Cur: REAL;
	i_iGrpUnitNum_Pu : INT;
	i_aiGrpUnitList: ARRAY [1..MAX_UNIT_NUM] OF INT;
	i_iGrpLinkageAxisNum_Pu: INT;
	i_aiGrpLinkageAxisList : ARRAY [1..MAX_UNIT_NUM] OF INT;
//	i_palrAxisMotionVel: POINTER TO ARRAY [1..MAX_UNIT_NUM] OF LREAL;(*轴速度*)
	i_paxFlag_PressDne: POINTER TO ARRAY [1..MAX_UNIT_NUM] OF BOOL;
	//增加加速度及加加速度输入只2026.4.11.153755
	i_rVel_A: REAL;//加速度
	i_rVel_Jerk: REAL;//加加速度；
	i_arAxisVelPrf_Coeff1: ARRAY [1..MAX_UNIT_NUM] OF REAL;
	i_arAxisVelPrf_Coeff2: ARRAY [1..MAX_UNIT_NUM] OF REAL;
	i_arAxisVelPrf_Coeff3: ARRAY [1..MAX_UNIT_NUM] OF REAL;
	i_xFlag_Accing: BOOL;
	i_xFlag_Decing: BOOL;
END_VAR
VAR_OUTPUT
	o_alrAxisPrfVel: ARRAY [1..MAX_UNIT_NUM] OF LREAL;
END_VAR
VAR
	iN: INT;
	iUnitId: INT;
	iPrevAxisId: INT;
	iPrevPressLinkageAxisId: INT;
	rAxisVelPrf_Coeff1: REAL;
	rAxisVelPrf_Coeff2: REAL;
	rAxisVelPrf_Coeff3: REAL;
 	rAxisVelPrf_Coeff: REAL;
	rCompensate_Vel: REAL;
	rTmp: REAL;
END_VAR

{IMPLEMENTATION}
(*按照所有轴输出*)
IF i_xEn THEN
	FOR iN:=1 TO i_iGrpUnitNum_Pu BY 1 DO
		iUnitId:= i_aiGrpUnitList[iN];
	//	pstStAxisParam:=ADR(i_pstStShmGlobalParam^.astStAxisParam[iAxisId]);
		IF in=1 THEN(*第一个轴为主速度*)
			o_alrAxisPrfVel[iUnitId]:= i_rVel_Cur;
		ELSE
			(*寻找前一个联动合压轴id*)
			iPrevPressLinkageAxisId:=
				KS_GetPrevPressLinkageAxisId(iUnitId,
					i_iGrpLinkageAxisNum_Pu,
					ADR(i_aiGrpLinkageAxisList[in]),
					i_paxFlag_PressDne);

			iPrevAxisId:= i_aiGrpUnitList[iN-1];
			IF iPrevPressLinkageAxisId<>-1 THEN(*找到了合压的前一个轴*)
				iPrevAxisId:=iPrevPressLinkageAxisId;
			ELSE;(*如果没找到，就用当前轴的前一个轴*)
			END_IF
			(*系数通过轴参数获取*)
			IF i_arAxisVelPrf_Coeff1[iUnitId]=0 THEN
				i_arAxisVelPrf_Coeff1[iUnitId]:= -200;
			END_IF
			rAxisVelPrf_Coeff1:=i_arAxisVelPrf_Coeff1[iUnitId];
			(*强制写为负值*)
			rAxisVelPrf_Coeff1:=-ABS(rAxisVelPrf_Coeff1);
			rAxisVelPrf_Coeff2:=i_arAxisVelPrf_Coeff2[iUnitId];
			rAxisVelPrf_Coeff3:=i_arAxisVelPrf_Coeff3[iUnitId];

			(*减加速度过程中修改加加速度的系数@2024.12.21.172422*)
			rAxisVelPrf_Coeff:=1;
			IF (i_rVel_Jerk<0 AND i_xFlag_Accing) OR
				(i_rVel_Jerk>0 AND i_xFlag_Decing) THEN
				rAxisVelPrf_Coeff:=rAxisVelPrf_Coeff3;
			END_IF

			(*前一个色组的速度基础上叠加补偿量@2024.12.29.134559*)
			(*补偿量*)
			rCompensate_Vel:=1/(rAxisVelPrf_Coeff1)*
						(i_rVel_Jerk*rAxisVelPrf_Coeff+rAxisVelPrf_Coeff2*i_rVel_A);

			rTmp:=rCompensate_Vel;

			o_alrAxisPrfVel[iUnitId]:=rTmp+o_alrAxisPrfVel[iPrevAxisId];
		END_IF
	END_FOR
END_IF

(* ---- KS_FB_GetAcceleToSync.st ---- *)
(*@CES
Name=KS_FB_GetAcceleToSync
Type=FunctionBlock
TypeGuid=6f9dac99-8de1-4efc-8465-68ac443b7d08
Guid=1e03253e-94af-4af4-b6f9-e65dddefd7f7
HasDeclaration=True
HasImplementation=True
*)
{DECLARATION}
FUNCTION_BLOCK KS_FB_GetAcceleToSync(*计算为了停止再开速度同步时位置同步的加速度*)
(*2022.11.29.232720 轴速度是带方向|计算取值需要增加取绝对值*)
VAR_INPUT
	i_xEn:BOOL;
	i_iGrpId: INT;
	i_iGrpAxisNum_Pu: INT; (*色组轴数量*)
	i_pstStSysParam: POINTER TO StSysParam;
//	i_pstStGrpParam: POINTER TO StGrpParam;(*系参数访问入口|*)
	i_paiGrpAxisList: POINTER TO ARRAY [1..MAX_UNIT_NUM] OF INT; (*系内所有轴的列表*)
//	i_pastStAxisParam: POINTER TO ARRAY [1..MAX_STATION_NUM] OF StAxisParam;
	i_pabyAxisMotionSts: POINTER TO ARRAY [1..MAX_STATION_NUM] OF BYTE;(*轴运动状态*)
	i_palrAcceleToSync:POINTER TO ARRAY [1..16] OF LREAL;(*同步加速度*)
	i_palrTimeToSync:POINTER TO ARRAY [1..16] OF LREAL;(*同步加到目标速度的时间*)
	i_palrRelatePos_Final:POINTER TO ARRAY [1..16,1..16] OF LREAL;(*做成16个轴|
													记录目标轴和当前轴的相对位置值|最后恢复的位置差
													一维下标为当前轴号，二维下标为目标轴号*)
	i_palrRelatePosToSync:POINTER TO ARRAY [1..16,1..16] OF LREAL;(*做成16个轴|
												记录目标轴和当前轴的相对位置值|开始切换到同步状态时的位置差
												一维下标为当前轴号，二维下标为目标轴号*)
	(*2022.7.17.165046 增加标志表征从同步状态退出到了其他状态|*)
END_VAR
VAR_OUTPUT
	o_xEn:BOOL;
END_VAR
VAR
	iN: INT;
	pstStUnitParam_Save: POINTER TO StUnitParam_Save;
	pstStUnitParam_UnSave: POINTER TO StUnitParam_UnSave;
	abyLastAxisMotionSts: ARRAY [1..MAX_STATION_NUM] OF BYTE;(*轴运动状态上个周期值*)
	iUnitId: INT;

	aiUnitId_Tar: ARRAY [1..16] OF INT;(*目标轴号|下标为当前轴号*)
	iUnitId_Tar: INT;
	alrVel_Sa: ARRAY [1..16] OF LREAL;(*起始速度*)
	alrVel_Tar: ARRAY [1..16] OF LREAL;(*目标速度*)
	lrTimeToSync:LREAL;(*去同步状态的时间|到达速度时位置同步*)
	axAxisMotionSts_0ToNot0:ARRAY [1..16] OF BOOL;(*轴状态从0切换到非0标志|用来防止开机时候有轴处于2
												状态-切换到5状态时候触发计算同步函数*)
END_VAR
{IMPLEMENTATION}
IF i_iGrpAxisNum_Pu>1 AND(*最少2个轴*)
	i_paiGrpAxisList<>0 AND
//	i_pastStAxisParam<>0 AND
	i_pabyAxisMotionSts<>0 AND
	i_pstStSysParam<>0 AND
	i_palrAcceleToSync<>0 AND
	i_palrTimeToSync<>0 AND
	i_palrRelatePos_Final<>0 AND
	i_palrRelatePosToSync<>0 THEN

	FOR iN:=1 TO i_iGrpAxisNum_Pu BY 1 DO
		iUnitId:=i_paiGrpAxisList^[iN];
		IF i_palrAcceleToSync<>0 THEN
			i_palrAcceleToSync^[iUnitId]:=0;
		END_IF
		IF i_palrTimeToSync<>0 THEN
			i_palrTimeToSync^[iUnitId]:=0;
		END_IF
	END_FOR

//	i_pastStAxisParam^[1].lrPT_Pos;
//	i_pastStAxisParam^[2].lrPT_Pos;

	IF i_xEn THEN(*使能*)
		FOR iN:=1 TO i_iGrpAxisNum_Pu BY 1 DO
			iUnitId:=i_paiGrpAxisList^[iN];
			pstStUnitParam_Save:=ADR(i_pstStSysParam^.astStUnitParam_Save[iUnitId]);
			pstStUnitParam_UnSave:=ADR(i_pstStSysParam^.astStUnitParam_UnSave[iUnitId]);
			IF iUnitId>0 AND iUnitId<=16 THEN
				(*从同步状态切换出去时记录位置偏差*)
				IF i_pabyAxisMotionSts^[iUnitId]<>0 AND
					abyLastAxisMotionSts[iUnitId]=0 THEN
						axAxisMotionSts_0ToNot0[iUnitId]:=TRUE;
						KS_GetRelatePos(
							iUnitId(*i_iAxisId_Cur*),
							i_iGrpAxisNum_Pu(*i_iGrpAxisNum_Pu*),
							i_paiGrpAxisList(*i_paiGrpAxisList*),
							ADR(i_pstStSysParam^.astStUnitParam_Save),(*i_pastStAxisParam*)
							ADR(i_pstStSysParam^.astStUnitParam_UnSave),(*i_pastStAxisParam*)
							ADR(i_palrRelatePos_Final^[iUnitId,1])(*i_palrRelatePos*));
				END_IF

				(*由其他状态进入同步运动时的位置偏差值*)
				IF i_pabyAxisMotionSts^[iUnitId]=5 AND
					abyLastAxisMotionSts[iUnitId]<>5 THEN
						KS_GetRelatePos(
							iUnitId(*i_iAxisId_Cur*),
							i_iGrpAxisNum_Pu(*i_iGrpAxisNum_Pu*),
							i_paiGrpAxisList(*i_paiGrpAxisList*),
							ADR(i_pstStSysParam^.astStUnitParam_Save),(*i_pastStAxisParam*)
							ADR(i_pstStSysParam^.astStUnitParam_UnSave),(*i_pastStAxisParam*)
							ADR(i_palrRelatePosToSync^[iUnitId,1])(*i_palrRelatePos*));

					(*记录当前速度和目标速度*)
					alrVel_Sa[iUnitId]:=ABS(pstStUnitParam_UnSave^.rAxisVel_PrnRoller);
					alrVel_Tar[iUnitId]:= i_pstStSysParam^.astStGrpParam_UnSave[i_iGrpId].rVel_Cur;

					(*寻找合适的目标轴号*)
					aiUnitId_Tar[iUnitId]:=
							KS_GetUnitId_Tar(
								iUnitId(*i_iAxisId_Cur*),
								i_iGrpAxisNum_Pu(*i_iGrpAxisNum_Pu*),
								i_paiGrpAxisList(*i_paiGrpAxisList*),
								ADR(i_pstStSysParam^.astStUnitParam_Save),(*i_pastStAxisParam*)
								ADR(i_pstStSysParam^.astStUnitParam_UnSave),(*i_pastStAxisParam*)
								i_pabyAxisMotionSts(*i_pabyAxisMotionSts*));

				ELSIF i_pabyAxisMotionSts^[iUnitId]<>5 THEN(*退出了加速到同步状态清除计算标志*)
					aiUnitId_Tar[iUnitId]:=-1;
				END_IF
			END_IF
		END_FOR

		(*计算当前轴的加速度*)
		FOR iN:=1 TO i_iGrpAxisNum_Pu BY 1 DO
			iUnitId:=i_paiGrpAxisList^[iN];
			pstStUnitParam_Save:=ADR(i_pstStSysParam^.astStUnitParam_Save[iUnitId]);
			pstStUnitParam_UnSave:=ADR(i_pstStSysParam^.astStUnitParam_UnSave[iUnitId]);
			(*计算当前轴加速到同步速度时的加速度*)
			lrTimeToSync:=0;
			IF iUnitId>0 AND iUnitId<=16 THEN
				iUnitId_Tar:=aiUnitId_Tar[iUnitId];
				IF iUnitId_Tar>0 AND iUnitId_Tar<=16 AND
					axAxisMotionSts_0ToNot0[iUnitId] THEN(*2022.7.17.165820 用来防止开机时候有轴处于2
																状态-切换到5状态时候触发计算同步函数*)
					lrTimeToSync:=KS_CalcMovePara(
										alrVel_Sa[iUnitId](*i_lrVelSa*),
										alrVel_Tar[iUnitId](*i_lrVelTar*),
										gc_iCycleTime_Motion(*i_iDeltime*),
										pstStUnitParam_Save^.rGirth_PrnRoller(*i_lrGirth_Axis*),
										UINT_TO_LREAL(pstStUnitParam_Save^.uiNum_PrnRoller)/pstStUnitParam_Save^.uiDen_PrnRoller(*i_lrReductionRatio*),
										i_palrRelatePosToSync^[iUnitId,iUnitId_Tar](*i_lrDeltPos_Init*),
										i_palrRelatePos_Final^[iUnitId,iUnitId_Tar](*i_lrDeltPos_Final*),
										LREAL_TO_DWORD(GC_LRMOTORPPR)(*i_dwMotorPPR*),
										10(*i_iSetTime*));
				END_IF

				IF i_palrTimeToSync<>0 THEN
					i_palrTimeToSync^[iUnitId]:=lrTimeToSync;
				END_IF
				IF lrTimeToSync>0 THEN
					IF i_palrAcceleToSync<>0 THEN
						i_palrAcceleToSync^[iUnitId]:=(alrVel_Tar[iUnitId]-alrVel_Sa[iUnitId])/lrTimeToSync/1000;
					END_IF
				END_IF
			END_IF
		END_FOR
	ELSE(*非使能*)
		SysMemSet(ADR(axAxisMotionSts_0ToNot0),0,SIZEOF(axAxisMotionSts_0ToNot0));
	END_IF
	o_xEn:=i_xEn;
ELSE
	o_xEn:=FALSE;
END_IF

(*备份状态值*)
IF i_iGrpAxisNum_Pu>1 AND(*最少2个轴*)
	i_paiGrpAxisList<>0 THEN
	FOR iN:=1 TO i_iGrpAxisNum_Pu BY 1 DO
		iUnitId:=i_paiGrpAxisList^[iN];
		abyLastAxisMotionSts[iUnitId]:=i_pabyAxisMotionSts^[iUnitId];
	END_FOR
END_IF
